// TIA Portal V20 export
// export: Created 2026-10-12T15:46:53.376981Z, ExportSetting WithDefaults, DisplayName Totally Integrated Automation Portal, DisplayVersion V20, DisplayName TIA Portal Openness, DisplayVersion V20, DisplayName TIA Portal Teamcenter Gateway, DisplayVersion V20, DisplayName TIA Portal Version Control Interface, DisplayVersion V20, DisplayName SINAMICS Startdrive Advanced, DisplayVersion V20 SP1 Update 2, DisplayName SINAMICS Startdrive G110M, G120, G120C, G120D, G120P, G115D, DisplayVersion V20 SP1 Update 2, DisplayName SINAMICS Startdrive G130, G150, S120, S150, SINAMICS MV, G220, S200, S210, DisplayVersion V20 SP1 Update 2, DisplayName STEP 7 Professional, DisplayVersion V20, DisplayName STEP 7 Safety, DisplayVersion V20, DisplayName WinCC Basic/Comfort/Advanced, DisplayVersion V20, DisplayName WinCC Professional, DisplayVersion V20, DisplayName WinCC Unified, DisplayVersion V20
FUNCTION "FRK_CfgSetWalk_InnerUnit" : Bool   // FC153, SCL
{ S7_Optimized_Access := 'TRUE' }
VERSION : 0.1
// stored: AutoNumber true, IsIECCheckEnabled false, SetENOAutomatically false, UDAEnableTagReadback false
   VAR_INPUT
      RootIndex : Int;
      Phase : Int;
      Access : "FRK_Access";
      Ready : Bool;
   END_VAR
   VAR_IN_OUT
      Module : "FB_InnerUnit";
   END_VAR
   VAR_TEMP
      Slot : Int;
      Stored : Int;
      Ok : Bool;
   END_VAR
BEGIN

   #FRK_CfgSetWalk_InnerUnit := FALSE;
   IF #Phase = 1 THEN
       #Module.ConfigStageParCfg := #Module.ParCfg;
   END_IF;
   IF #Phase = 1 THEN
       #Module.ConfigStageStationCfg := #Module.StationCfg;
   END_IF;
   IF "FRK_SetRuntime".Work[#RootIndex].Payload.Info.Kind = 0 THEN
       "FRK_CfgDef_InnerUnit"(FieldIndex := 1);
       "FRK_SetRuntime".Work[#RootIndex].RejectScope := #Module.Status.Name;
       "FRK_SetRuntime".Work[#RootIndex].RejectKey := "FRK_ConfigScratch".Entry.WriteKey;
       IF #Phase = 0 THEN
           IF #Access.CurrentLevel < MAX(IN1 := #Access.Policy.Required[0], IN2 := "FRK_ConfigScratch".MinRead) THEN
               RETURN;
           END_IF;
           #Ok := "FRK_ConfigGet"(Scope := #Module.Status.Name, ModelCode := "FRK_SetRuntime".Work[#RootIndex].Payload.Info.ModelCode);
           IF NOT #Ok OR "FRK_SetRuntime".Work[#RootIndex].Payload.Info.RecordCount >= 24 THEN
               RETURN;
           END_IF;
           #Slot := "FRK_SetRuntime".Work[#RootIndex].Payload.Info.RecordCount + 1;
           "FRK_SetRuntime".Work[#RootIndex].Payload.Records[#Slot].Scope := #Module.Status.Name;
           "FRK_SetRuntime".Work[#RootIndex].Payload.Records[#Slot].WriteKey := "FRK_ConfigScratch".Entry.WriteKey;
           "FRK_SetRuntime".Work[#RootIndex].Payload.Records[#Slot].Revision := "FRK_ConfigScratch".Entry.WriteRevision;
           "FRK_SetRuntime".Work[#RootIndex].Payload.Records[#Slot].Kind := "FRK_ConfigScratch".Entry.ConfigKind;
           "FRK_SetRuntime".Work[#RootIndex].Payload.Records[#Slot].ValueType := "FRK_ConfigScratch".Entry.ValueType;
           "FRK_SetRuntime".Work[#RootIndex].Payload.Records[#Slot].ValueText := WSTRING_TO_STRING("FRK_ConfigScratch".Entry.ValueText);
           "FRK_SetRuntime".Work[#RootIndex].Payload.Info.RecordCount := #Slot;
       ELSIF #Phase = 2 THEN
           #Slot := "FRK_SetRecord"(RootIndex := #RootIndex, Scope := #Module.Status.Name, WriteKey := "FRK_ConfigScratch".Entry.WriteKey);
           #Stored := "FRK_ConfigFind"(Scope := #Module.Status.Name, Key := "FRK_ConfigScratch".Entry.WriteKey, ModelCode := "FRK_SetRuntime".Work[#RootIndex].Payload.Info.ModelCode);
           "FRK_ConfigStore".Rows[#Stored].Record := "FRK_SetRuntime".Work[#RootIndex].Payload.Records[#Slot];
           "FRK_ConfigStore".Rows[#Stored].SchemaVersion := "FRK_ConfigScratch".Schema;
       ELSE
           #Slot := "FRK_SetCheck"(RootIndex := #RootIndex, Scope := #Module.Status.Name, Access := #Access, Ready := #Ready, WriteAccess := #Phase <> 3);
           IF #Slot = 0 THEN
               RETURN;
           END_IF;
           IF #Phase = 1 THEN
               #Module.ConfigStageParCfg.Timeout := DINT_TO_TIME(LINT_TO_DINT("FRK_ConfigScratch".Value.Number));
           END_IF;
       END_IF;
   END_IF;
   IF "FRK_SetRuntime".Work[#RootIndex].Payload.Info.Kind = 0 THEN
       "FRK_CfgDef_InnerUnit"(FieldIndex := 2);
       "FRK_SetRuntime".Work[#RootIndex].RejectScope := #Module.Status.Name;
       "FRK_SetRuntime".Work[#RootIndex].RejectKey := "FRK_ConfigScratch".Entry.WriteKey;
       IF #Phase = 0 THEN
           IF #Access.CurrentLevel < MAX(IN1 := #Access.Policy.Required[0], IN2 := "FRK_ConfigScratch".MinRead) THEN
               RETURN;
           END_IF;
           #Ok := "FRK_ConfigGet"(Scope := #Module.Status.Name, ModelCode := "FRK_SetRuntime".Work[#RootIndex].Payload.Info.ModelCode);
           IF NOT #Ok OR "FRK_SetRuntime".Work[#RootIndex].Payload.Info.RecordCount >= 24 THEN
               RETURN;
           END_IF;
           #Slot := "FRK_SetRuntime".Work[#RootIndex].Payload.Info.RecordCount + 1;
           "FRK_SetRuntime".Work[#RootIndex].Payload.Records[#Slot].Scope := #Module.Status.Name;
           "FRK_SetRuntime".Work[#RootIndex].Payload.Records[#Slot].WriteKey := "FRK_ConfigScratch".Entry.WriteKey;
           "FRK_SetRuntime".Work[#RootIndex].Payload.Records[#Slot].Revision := "FRK_ConfigScratch".Entry.WriteRevision;
           "FRK_SetRuntime".Work[#RootIndex].Payload.Records[#Slot].Kind := "FRK_ConfigScratch".Entry.ConfigKind;
           "FRK_SetRuntime".Work[#RootIndex].Payload.Records[#Slot].ValueType := "FRK_ConfigScratch".Entry.ValueType;
           "FRK_SetRuntime".Work[#RootIndex].Payload.Records[#Slot].ValueText := WSTRING_TO_STRING("FRK_ConfigScratch".Entry.ValueText);
           "FRK_SetRuntime".Work[#RootIndex].Payload.Info.RecordCount := #Slot;
       ELSIF #Phase = 2 THEN
           #Slot := "FRK_SetRecord"(RootIndex := #RootIndex, Scope := #Module.Status.Name, WriteKey := "FRK_ConfigScratch".Entry.WriteKey);
           #Stored := "FRK_ConfigFind"(Scope := #Module.Status.Name, Key := "FRK_ConfigScratch".Entry.WriteKey, ModelCode := "FRK_SetRuntime".Work[#RootIndex].Payload.Info.ModelCode);
           "FRK_ConfigStore".Rows[#Stored].Record := "FRK_SetRuntime".Work[#RootIndex].Payload.Records[#Slot];
           "FRK_ConfigStore".Rows[#Stored].SchemaVersion := "FRK_ConfigScratch".Schema;
       ELSE
           #Slot := "FRK_SetCheck"(RootIndex := #RootIndex, Scope := #Module.Status.Name, Access := #Access, Ready := #Ready, WriteAccess := #Phase <> 3);
           IF #Slot = 0 THEN
               RETURN;
           END_IF;
           IF #Phase = 1 THEN
               #Module.ConfigStageParCfg.Preset := LINT_TO_DINT("FRK_ConfigScratch".Value.Number);
           END_IF;
       END_IF;
   END_IF;
   IF "FRK_SetRuntime".Work[#RootIndex].Payload.Info.Kind = 1 THEN
       "FRK_CfgDef_InnerUnit"(FieldIndex := 3);
       "FRK_SetRuntime".Work[#RootIndex].RejectScope := #Module.Status.Name;
       "FRK_SetRuntime".Work[#RootIndex].RejectKey := "FRK_ConfigScratch".Entry.WriteKey;
       IF #Phase = 0 THEN
           IF #Access.CurrentLevel < MAX(IN1 := #Access.Policy.Required[0], IN2 := "FRK_ConfigScratch".MinRead) THEN
               RETURN;
           END_IF;
           #Ok := "FRK_ConfigGet"(Scope := #Module.Status.Name, ModelCode := "FRK_SetRuntime".Work[#RootIndex].Payload.Info.ModelCode);
           IF NOT #Ok OR "FRK_SetRuntime".Work[#RootIndex].Payload.Info.RecordCount >= 24 THEN
               RETURN;
           END_IF;
           #Slot := "FRK_SetRuntime".Work[#RootIndex].Payload.Info.RecordCount + 1;
           "FRK_SetRuntime".Work[#RootIndex].Payload.Records[#Slot].Scope := #Module.Status.Name;
           "FRK_SetRuntime".Work[#RootIndex].Payload.Records[#Slot].WriteKey := "FRK_ConfigScratch".Entry.WriteKey;
           "FRK_SetRuntime".Work[#RootIndex].Payload.Records[#Slot].Revision := "FRK_ConfigScratch".Entry.WriteRevision;
           "FRK_SetRuntime".Work[#RootIndex].Payload.Records[#Slot].Kind := "FRK_ConfigScratch".Entry.ConfigKind;
           "FRK_SetRuntime".Work[#RootIndex].Payload.Records[#Slot].ValueType := "FRK_ConfigScratch".Entry.ValueType;
           "FRK_SetRuntime".Work[#RootIndex].Payload.Records[#Slot].ValueText := WSTRING_TO_STRING("FRK_ConfigScratch".Entry.ValueText);
           "FRK_SetRuntime".Work[#RootIndex].Payload.Info.RecordCount := #Slot;
       ELSIF #Phase = 2 THEN
           #Slot := "FRK_SetRecord"(RootIndex := #RootIndex, Scope := #Module.Status.Name, WriteKey := "FRK_ConfigScratch".Entry.WriteKey);
           #Stored := "FRK_ConfigFind"(Scope := #Module.Status.Name, Key := "FRK_ConfigScratch".Entry.WriteKey, ModelCode := "FRK_SetRuntime".Work[#RootIndex].Payload.Info.ModelCode);
           "FRK_ConfigStore".Rows[#Stored].Record := "FRK_SetRuntime".Work[#RootIndex].Payload.Records[#Slot];
           "FRK_ConfigStore".Rows[#Stored].SchemaVersion := "FRK_ConfigScratch".Schema;
       ELSE
           #Slot := "FRK_SetCheck"(RootIndex := #RootIndex, Scope := #Module.Status.Name, Access := #Access, Ready := #Ready, WriteAccess := #Phase <> 3);
           IF #Slot = 0 THEN
               RETURN;
           END_IF;
           IF #Phase = 1 THEN
               #Module.ConfigStageStationCfg.SiteLabel := "FRK_ConfigScratch".Value.Text;
           END_IF;
       END_IF;
   END_IF;
   IF "FRK_SetRuntime".Work[#RootIndex].Payload.Info.Kind = 1 THEN
       "FRK_CfgDef_InnerUnit"(FieldIndex := 4);
       "FRK_SetRuntime".Work[#RootIndex].RejectScope := #Module.Status.Name;
       "FRK_SetRuntime".Work[#RootIndex].RejectKey := "FRK_ConfigScratch".Entry.WriteKey;
       IF #Phase = 0 THEN
           IF #Access.CurrentLevel < MAX(IN1 := #Access.Policy.Required[0], IN2 := "FRK_ConfigScratch".MinRead) THEN
               RETURN;
           END_IF;
           #Ok := "FRK_ConfigGet"(Scope := #Module.Status.Name, ModelCode := "FRK_SetRuntime".Work[#RootIndex].Payload.Info.ModelCode);
           IF NOT #Ok OR "FRK_SetRuntime".Work[#RootIndex].Payload.Info.RecordCount >= 24 THEN
               RETURN;
           END_IF;
           #Slot := "FRK_SetRuntime".Work[#RootIndex].Payload.Info.RecordCount + 1;
           "FRK_SetRuntime".Work[#RootIndex].Payload.Records[#Slot].Scope := #Module.Status.Name;
           "FRK_SetRuntime".Work[#RootIndex].Payload.Records[#Slot].WriteKey := "FRK_ConfigScratch".Entry.WriteKey;
           "FRK_SetRuntime".Work[#RootIndex].Payload.Records[#Slot].Revision := "FRK_ConfigScratch".Entry.WriteRevision;
           "FRK_SetRuntime".Work[#RootIndex].Payload.Records[#Slot].Kind := "FRK_ConfigScratch".Entry.ConfigKind;
           "FRK_SetRuntime".Work[#RootIndex].Payload.Records[#Slot].ValueType := "FRK_ConfigScratch".Entry.ValueType;
           "FRK_SetRuntime".Work[#RootIndex].Payload.Records[#Slot].ValueText := WSTRING_TO_STRING("FRK_ConfigScratch".Entry.ValueText);
           "FRK_SetRuntime".Work[#RootIndex].Payload.Info.RecordCount := #Slot;
       ELSIF #Phase = 2 THEN
           #Slot := "FRK_SetRecord"(RootIndex := #RootIndex, Scope := #Module.Status.Name, WriteKey := "FRK_ConfigScratch".Entry.WriteKey);
           #Stored := "FRK_ConfigFind"(Scope := #Module.Status.Name, Key := "FRK_ConfigScratch".Entry.WriteKey, ModelCode := "FRK_SetRuntime".Work[#RootIndex].Payload.Info.ModelCode);
           "FRK_ConfigStore".Rows[#Stored].Record := "FRK_SetRuntime".Work[#RootIndex].Payload.Records[#Slot];
           "FRK_ConfigStore".Rows[#Stored].SchemaVersion := "FRK_ConfigScratch".Schema;
       ELSE
           #Slot := "FRK_SetCheck"(RootIndex := #RootIndex, Scope := #Module.Status.Name, Access := #Access, Ready := #Ready, WriteAccess := #Phase <> 3);
           IF #Slot = 0 THEN
               RETURN;
           END_IF;
           IF #Phase = 1 THEN
               #Module.ConfigStageStationCfg.LongText := "FRK_ConfigScratch".Value.Text;
           END_IF;
       END_IF;
   END_IF;
   IF "FRK_SetRuntime".Work[#RootIndex].Payload.Info.Kind = 1 THEN
       "FRK_CfgDef_InnerUnit"(FieldIndex := 5);
       "FRK_SetRuntime".Work[#RootIndex].RejectScope := #Module.Status.Name;
       "FRK_SetRuntime".Work[#RootIndex].RejectKey := "FRK_ConfigScratch".Entry.WriteKey;
       IF #Phase = 0 THEN
           IF #Access.CurrentLevel < MAX(IN1 := #Access.Policy.Required[0], IN2 := "FRK_ConfigScratch".MinRead) THEN
               RETURN;
           END_IF;
           #Ok := "FRK_ConfigGet"(Scope := #Module.Status.Name, ModelCode := "FRK_SetRuntime".Work[#RootIndex].Payload.Info.ModelCode);
           IF NOT #Ok OR "FRK_SetRuntime".Work[#RootIndex].Payload.Info.RecordCount >= 24 THEN
               RETURN;
           END_IF;
           #Slot := "FRK_SetRuntime".Work[#RootIndex].Payload.Info.RecordCount + 1;
           "FRK_SetRuntime".Work[#RootIndex].Payload.Records[#Slot].Scope := #Module.Status.Name;
           "FRK_SetRuntime".Work[#RootIndex].Payload.Records[#Slot].WriteKey := "FRK_ConfigScratch".Entry.WriteKey;
           "FRK_SetRuntime".Work[#RootIndex].Payload.Records[#Slot].Revision := "FRK_ConfigScratch".Entry.WriteRevision;
           "FRK_SetRuntime".Work[#RootIndex].Payload.Records[#Slot].Kind := "FRK_ConfigScratch".Entry.ConfigKind;
           "FRK_SetRuntime".Work[#RootIndex].Payload.Records[#Slot].ValueType := "FRK_ConfigScratch".Entry.ValueType;
           "FRK_SetRuntime".Work[#RootIndex].Payload.Records[#Slot].ValueText := WSTRING_TO_STRING("FRK_ConfigScratch".Entry.ValueText);
           "FRK_SetRuntime".Work[#RootIndex].Payload.Info.RecordCount := #Slot;
       ELSIF #Phase = 2 THEN
           #Slot := "FRK_SetRecord"(RootIndex := #RootIndex, Scope := #Module.Status.Name, WriteKey := "FRK_ConfigScratch".Entry.WriteKey);
           #Stored := "FRK_ConfigFind"(Scope := #Module.Status.Name, Key := "FRK_ConfigScratch".Entry.WriteKey, ModelCode := "FRK_SetRuntime".Work[#RootIndex].Payload.Info.ModelCode);
           "FRK_ConfigStore".Rows[#Stored].Record := "FRK_SetRuntime".Work[#RootIndex].Payload.Records[#Slot];
           "FRK_ConfigStore".Rows[#Stored].SchemaVersion := "FRK_ConfigScratch".Schema;
       ELSE
           #Slot := "FRK_SetCheck"(RootIndex := #RootIndex, Scope := #Module.Status.Name, Access := #Access, Ready := #Ready, WriteAccess := #Phase <> 3);
           IF #Slot = 0 THEN
               RETURN;
           END_IF;
           IF #Phase = 1 THEN
               #Module.ConfigStageStationCfg.Enabled := "FRK_ConfigScratch".Value.Flag;
           END_IF;
       END_IF;
   END_IF;
   IF #Phase = 2 AND "FRK_SetRuntime".Work[#RootIndex].Payload.Info.Kind = 0 THEN
       #Module.ParCfg := #Module.ConfigStageParCfg;
   END_IF;
   IF #Phase = 2 AND "FRK_SetRuntime".Work[#RootIndex].Payload.Info.Kind = 1 THEN
       #Module.StationCfg := #Module.ConfigStageStationCfg;
   END_IF;
   #Ok := "FRK_CfgSetWalk_DeclarationCell"(Module := #Module.Cell, RootIndex := #RootIndex, Phase := #Phase, Access := #Access, Ready := #Ready);
   IF NOT #Ok THEN
       RETURN;
   END_IF;
   #FRK_CfgSetWalk_InnerUnit := TRUE;
END_FUNCTION
